(* PLC project Vn_ctu_call, Beckhoff Automation GmbH TwinCAT PLC Control 3.5.13.21 *)
(* stored: creationDateTime 1970-01-01T00:00:00 *)

PROGRAM Vn_ctu_call

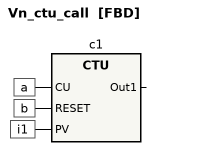
(* FBD diagram, written out as Structured Text *)
c1(CU := a, RESET := b, PV := i1);
END_PROGRAM
